TYPE ET_CfgAxisInExt3DGroup :
(
	ET_CfgAxisInExt3DGrp_eWaitExecute := 0,
	ET_CfgAxisInExt3DGrp_eReadExt3DAxisIds := 5,
	ET_CfgAxisInExt3DGrp_eDone := 197,
	ET_CfgAxisInExt3DGrp_eError := 198,
	ET_CfgAxisInExt3DGrp_eNoExecute := 199
);
END_TYPE

(* stored: Version 1.1.0.1, ProductVersion 3.1.4024.15
   DUT ET_CfgAxisInExt3DGroup: Id {59a689a1-e9b9-42ee-b459-eec819f00c1d} *)
